(* Generated by scripts/make_testbench.py. Do not edit.
   OB1 of the test project: one call of the bench per cycle; the result is copied to DB_TestResult. *)
ORGANIZATION_BLOCK "Main"
TITLE = "Main Program Sweep (Cycle)"
{ S7_Optimized_Access := 'TRUE' }
VERSION : 0.1
   VAR_TEMP
      bits : DWord;
   END_VAR
BEGIN
  "TB_BENCH_DB"(enable := TRUE,
                Done => "DB_TestResult".Done,
                CasesTotal => "DB_TestResult".CasesTotal,
                CasesRun => "DB_TestResult".CasesRun,
                CasesPassed => "DB_TestResult".CasesPassed,
                CasesFailed => "DB_TestResult".CasesFailed,
                FirstFailedCase => "DB_TestResult".FirstFailedCase,
                FirstFailedCheck => "DB_TestResult".FirstFailedCheck,
                CasePassBits => #bits);
  "DB_TestResult".CasePassed[1] := (#bits AND DW#16#1) <> DW#16#0;
  "DB_TestResult".CasePassed[2] := (#bits AND DW#16#2) <> DW#16#0;
  "DB_TestResult".CasePassed[3] := (#bits AND DW#16#4) <> DW#16#0;
  "DB_TestResult".CasePassed[4] := (#bits AND DW#16#8) <> DW#16#0;
  "DB_TestResult".CasePassed[5] := (#bits AND DW#16#10) <> DW#16#0;
  "DB_TestResult".CasePassed[6] := (#bits AND DW#16#20) <> DW#16#0;
  "DB_TestResult".CasePassed[7] := (#bits AND DW#16#40) <> DW#16#0;
END_ORGANIZATION_BLOCK
